TYPE "ST_DeclarationOutImm"
VERSION : 0.1
   STRUCT
      "Sample" : DInt;
      "InitCount" : DInt;
      "StartCount" : DInt;
      "CyclicCount" : DInt;
      "AbortCount" : DInt;
      "ErrorAbortCount" : DInt;
      "DispatchCount" : DInt;
      "SeenValue" : DInt;
      "Ordered" : Bool;
      "Output" : Bool;
   END_STRUCT;
END_TYPE
